// TIA Portal V20 export
FUNCTION "POS3_0_Bausteinaufrufe" : Void   // FC27, STL
{ S7_Optimized_Access := 'TRUE' }
BEGIN

NETWORK
TITLE = 

      CALL  "POS3_0_Betriebsart";

      CALL  "POS3_0_Antriebe", "POS3_0_Antriebe_DB";

      CALL  "POS3_0_Melden_Visu", "POS3_0_Melden_Visu_DB";
      CALL  "POS3_0_Teileauswertung";

      CALL  "POS3_0_Messtechnik", "POS3_0_Messtechnik_DB";




NETWORK
TITLE = 

      A     "03_Betriebsart_DB".ACK_Taste;
      =     "POS3_0_Signal".Schrittkette.ACK_EF;



      CALL  "POS3_0_SK_Ablauf", "POS3_0_SK_Ablauf_DB"
      ( OFF_SQ         := "POS3_0_Signal".Schrittkette.OFF_SQ,
        INIT_SQ        := "POS3_0_Signal".Schrittkette.INIT_SQ,
        ACK_EF         := "POS3_0_Signal".Schrittkette.ACK_EF,
        REG_EF         := ,
        ACK_S          := ,
        REG_S          := ,
        HALT_SQ        := "POS3_0_Signal".Schrittkette.HALT_SQ,
        HALT_TM        := "POS3_0_Signal".Schrittkette.HALT_TM,
        ZERO_OP        := "POS3_0_Signal".Schrittkette.ZERO_OP,
        EN_IL          := "POS3_0_Signal".Schrittkette.EN_IL,
        EN_SV          := "POS3_0_Signal".Schrittkette.EN_SV,
        EN_ACKREQ      := ,
        EN_SSKIP       := ,
        DISP_SACT      := ,
        DISP_SEF       := ,
        DISP_SALL      := ,
        S_PREV         := "POS3_0_Signal".Schrittkette.S_PREV,
        S_NEXT         := "POS3_0_Signal".Schrittkette.S_NEXT,
        SW_AUTO        := "POS3_0_Signal".Schrittkette.SW_AUTO,
        SW_TAP         := "POS3_0_Signal".Schrittkette.SW_TAP,
        SW_TOP         := 0,
        SW_MAN         := "POS3_0_Signal".Schrittkette.SW_MAN,
        S_SEL          := "POS3_0_Signal".Schrittkette.S_SEL,
        S_SELOK        := ,
        S_ON           := "POS3_0_Signal".Schrittkette.S_ON,
        S_OFF          := "POS3_0_Signal".Schrittkette.S_OFF,
        T_PREV         := ,
        T_NEXT         := ,
        T_PUSH         := "POS3_0_Signal".Schrittkette.T_PUSH,
        EN_LMODE       := ,
        S_NO           := "POS3_0_Signal".Schrittkette.S_NO,
        S_MORE         := "POS3_0_Signal".Schrittkette.S_MORE,
        S_ACTIVE       := "POS3_0_Signal".Schrittkette.S_ACTIVE,
        S_TIME         := ,
        S_TIMEOK       := ,
        S_CRITLOC      := ,
        S_CRITLOCERR   := ,
        S_STATE        := ,
        T_NO           := ,
        T_MORE         := ,
        T_CRIT         := ,
        T_CRITOLD      := ,
        T_CRITFLT      := ,
        ERROR          := ,
        FAULT          := ,
        ERR_FLT        := "POS3_0_Signal".Schrittkette.ERR_FLT,
        SQ_ISOFF       := ,
        SQ_HALTED      := "POS3_0_Signal".Schrittkette.SQ_HALTED,
        TM_HALTED      := "POS3_0_Signal".Schrittkette.TM_HALTED,
        OP_ZEROED      := "POS3_0_Signal".Schrittkette.OP_ZEROED,
        IL_ENABLED     := "POS3_0_Signal".Schrittkette.IL_ENABELD,
        SV_ENABLED     := "POS3_0_Signal".Schrittkette.SV_ENABELD,
        ACKREQ_ENABLED := ,
        SSKIP_ENABLED  := ,
        SACT_DISP      := ,
        SEF_DISP       := ,
        SALL_DISP      := ,
        AUTO_ON        := "POS3_0_Signal".Schrittkette.AUTO_ON,
        TAP_ON         := "POS3_0_Signal".Schrittkette.TAP_ON,
        TOP_ON         := ,
        MAN_ON         := "POS3_0_Signal".Schrittkette.MAN_ON,
        LMODE_ENABLED  := 
      );


END_FUNCTION
